VAR_GLOBAL
    bButton : BOOL;
    bLightRelay : BOOL;
END_VAR

(* stored: Version 1.1.0.1
   GVL GVL_WorkshopSimulation: Id {45436E6A-4F26-4402-B386-C69AEFB90D94} *)
